(* IEC 61131-3 sources: plc-hackathon-2026/deliver/ME_v3_src (part 2) *)

(* ---- Team_Results.st ---- *)
// Team_Results: YEARLY totals checked by the jury against SimScore.total (tolerance 0.1 %).
// Energies [kWh] and costs [EUR], all LREAL. Updated every simulation step (interval k-1).
VAR_GLOBAL
	E_fne : LREAL;                      // PV production after curtailment
	E_fec : LREAL;                      // fixed consumption
	E_bess_chg : LREAL;                 // battery charge, bus side
	E_bess_dch : LREAL;                 // battery discharge, bus side
	E_ev : LREAL;                       // EV chargers total, bus side
	E_import : LREAL;                   // grid import
	E_export : LREAL;                   // grid export
	E_ev_ch : ARRAY[0..3] OF LREAL;     // per EV charger, bus side
	P_peak : LREAL;                     // [kW] highest monthly peak of the year (info)
	// cost components (spec 4.3)
	C_purchase : LREAL;                 // energy purchase
	C_revenue : LREAL;                  // export revenue (0.9 * price)
	C_grid : LREAL;                     // grid fee
	C_peak : LREAL;                     // peak power cost = sum of 12 monthly values
	C_total : LREAL;                    // purchase - revenue + grid + peak
	// same quantities with the simulator's SimScore.total names
	cost_energy : LREAL;                // purchase - revenue
	cost_grid : LREAL;
	cost_peak : LREAL;
	cost_total : LREAL;
	nLogged : DINT;                     // number of 15-min intervals logged (35040 after the final call)
END_VAR

(* ---- F_AlarmPush.st ---- *)
FUNCTION F_AlarmPush : BOOL
// Push a message into the alarm history (Team_HMI.aAlarmHist, newest at index 0), stamped with simulated time.
VAR_INPUT
	k : DINT;
	sStamp : STRING(20);
	iCode : INT;
	sText : STRING(80);
END_VAR
VAR
	i : INT;
END_VAR
// ---IMPL---
FOR i := 49 TO 1 BY -1 DO
	Team_HMI.aAlarmHist[i] := Team_HMI.aAlarmHist[i - 1];
END_FOR;
Team_HMI.aAlarmHist[0].k := k;
Team_HMI.aAlarmHist[0].sStamp := sStamp;
Team_HMI.aAlarmHist[0].iCode := iCode;
Team_HMI.aAlarmHist[0].sText := sText;
Team_HMI.nAlarms := Team_HMI.nAlarms + 1;
Team_HMI.sLastAlarm := sText;
F_AlarmPush := TRUE;

(* ---- F_BessMaxChg.st ---- *)
FUNCTION F_BessMaxChg : REAL
// Largest bus-side charge power [kW] the simulator accepts at this SoC (same clamp as Sim_Core).
VAR_INPUT
	rSoc : REAL;            // [%] SoC at start of the interval
END_VAR
// ---IMPL---
F_BessMaxChg := LREAL_TO_REAL(MAX(0.0, MIN(REAL_TO_LREAL(SimParam.BESS_MAX_CHG),
	(REAL_TO_LREAL(SimParam.BESS_SOC_MAX) - REAL_TO_LREAL(rSoc)) / 100.0 * REAL_TO_LREAL(SimParam.BESS_CAPACITY)
	/ (REAL_TO_LREAL(SimParam.TS_H) * REAL_TO_LREAL(SimParam.BESS_ETA_CHG)))));

(* ---- F_BessMaxDch.st ---- *)
FUNCTION F_BessMaxDch : REAL
// Largest bus-side discharge power [kW] the simulator accepts at this SoC (same clamp as Sim_Core).
VAR_INPUT
	rSoc : REAL;            // [%] SoC at start of the interval
END_VAR
// ---IMPL---
F_BessMaxDch := LREAL_TO_REAL(MAX(0.0, MIN(REAL_TO_LREAL(SimParam.BESS_MAX_DCH),
	(REAL_TO_LREAL(rSoc) - REAL_TO_LREAL(SimParam.BESS_SOC_MIN)) / 100.0 * REAL_TO_LREAL(SimParam.BESS_CAPACITY)
	* REAL_TO_LREAL(SimParam.BESS_ETA_DCH) / REAL_TO_LREAL(SimParam.TS_H))));

(* ---- F_DayType.st ---- *)
FUNCTION F_DayType : INT
// Day type for load forecasting: 0 = Monday..Friday, 1 = Saturday, 2 = Sunday.
VAR_INPUT
	iWeekday : INT;                     // 1 = Monday .. 7 = Sunday
END_VAR
// ---IMPL---
IF iWeekday = 6 THEN
	F_DayType := 1;
ELSIF iWeekday = 7 THEN
	F_DayType := 2;
ELSE
	F_DayType := 0;
END_IF;

(* ---- F_DtString.st ---- *)
FUNCTION F_DtString : STRING(20)
// DT -> "DD.MM.YYYY HH:MM" (simulated time). Pure calendar arithmetic, no clock access.
VAR_INPUT
	dtIn : DT;
END_VAR
VAR
	udSec : UDINT;
	iDoy : INT;
	iYear : INT;
	iMon : INT;
	iDim : INT;
	xLeap : BOOL;
	uH : USINT;
	uM : USINT;
END_VAR
// ---IMPL---
udSec := DT_TO_UDINT(dtIn);                          // seconds since 1970-01-01
uH := UDINT_TO_USINT((udSec MOD 86400) / 3600);
uM := UDINT_TO_USINT((udSec MOD 3600) / 60);
iDoy := UDINT_TO_INT(udSec / 86400);
iYear := 1970;
xLeap := FALSE;
WHILE iYear < 2200 DO
	xLeap := ((iYear MOD 4) = 0 AND (iYear MOD 100) <> 0) OR ((iYear MOD 400) = 0);
	IF xLeap THEN iDim := 366; ELSE iDim := 365; END_IF;
	IF iDoy < iDim THEN EXIT; END_IF;
	iDoy := iDoy - iDim;
	iYear := iYear + 1;
END_WHILE;
iMon := 1;
WHILE iMon < 12 DO
	CASE iMon OF
		2: IF xLeap THEN iDim := 29; ELSE iDim := 28; END_IF;
		4, 6, 9, 11: iDim := 30;
	ELSE
		iDim := 31;
	END_CASE;
	IF iDoy < iDim THEN EXIT; END_IF;
	iDoy := iDoy - iDim;
	iMon := iMon + 1;
END_WHILE;
F_DtString := CONCAT(CONCAT(CONCAT(F_Pad2(INT_TO_USINT(iDoy + 1)), '.'), CONCAT(F_Pad2(INT_TO_USINT(iMon)), '.')),
	CONCAT(CONCAT(INT_TO_STRING(iYear), ' '), CONCAT(CONCAT(F_Pad2(uH), ':'), F_Pad2(uM))));

(* ---- F_EnergyPrice.st ---- *)
FUNCTION F_EnergyPrice : REAL
// Energy price [EUR/kWh] of interval k for the selected price model (same series the simulator uses).
//   iMode 0 = two-tariff Elektra (per calendar quarter, VT/NT), 1 = day-ahead (Team_Prices.aDA)
VAR_INPUT
	k : DINT;               // interval 0..35039
	iMonth : INT;           // 1..12 of interval k
	xHigh : BOOL;           // VT of interval k (t_sim.tariff_high)
	iMode : INT;            // SimCtrl.price_mode
END_VAR
VAR
	iQ : INT;
END_VAR
// ---IMPL---
IF iMode = 1 THEN
	F_EnergyPrice := Team_Prices.aDA[LIMIT(0, k, 35039)];
ELSE
	iQ := LIMIT(1, (iMonth - 1) / 3 + 1, 4);
	IF xHigh THEN
		F_EnergyPrice := Team_Prices.TT_VT[iQ];
	ELSE
		F_EnergyPrice := Team_Prices.TT_NT[iQ];
	END_IF;
END_IF;

(* ---- F_Pad2.st ---- *)
FUNCTION F_Pad2 : STRING(2)
// Two-digit zero padded number for date/time strings.
VAR_INPUT
	v : USINT;
END_VAR
// ---IMPL---
IF v < 10 THEN
	F_Pad2 := CONCAT('0', USINT_TO_STRING(v));
ELSE
	F_Pad2 := USINT_TO_STRING(v);
END_IF;

(* ---- F_PeakCap.st ---- *)
FUNCTION F_PeakCap : REAL
// Lowest monthly import cap [kW] the battery can hold over the horizon for the given net-load
// forecast (bisection). The battery covers load above the cap and recharges below it.
// Never below rFloor (the peak already paid this month), never above rLimImp.
VAR_INPUT
	h : INT;                            // horizon length
	rE0 : REAL;                         // usable stored energy now [kWh]
	rFloor : REAL;                      // peak already reached this month [kW]
	rLimImp : REAL;                     // import limit [kW]
END_VAR
VAR_IN_OUT
	aLoad : ARRAY[0..191] OF REAL;      // net-load forecast [kW]
END_VAR
VAR
	n : INT;
	i : INT;
	rMid : REAL;
	rLo : REAL;
	rHi : REAL;
	rE : REAL;
	rG : REAL;
	rNeed : REAL;
	rEuse : REAL;
	xOk : BOOL;
END_VAR
// ---IMPL---
rEuse := (SimParam.BESS_SOC_MAX - SimParam.BESS_SOC_MIN) / 100.0 * SimParam.BESS_CAPACITY;
F_PeakCap := rFloor;
rLo := rFloor;
rHi := rLimImp;
FOR n := 0 TO 12 DO
	IF n = 0 THEN
		rMid := rFloor;
	ELSE
		rMid := 0.5 * (rLo + rHi);
	END_IF;
	xOk := TRUE;
	rE := rE0;
	FOR i := 0 TO h - 1 DO
		rG := aLoad[i];
		IF rG > rMid THEN
			rNeed := rG - rMid;
			rE := rE - rNeed * SimParam.TS_H / SimParam.BESS_ETA_DCH;
			IF rNeed > SimParam.BESS_MAX_DCH OR rE < 0.0 THEN
				xOk := FALSE;
				EXIT;
			END_IF;
		ELSE
			rE := rE + MIN(MIN(rMid - rG, SimParam.BESS_MAX_CHG), (rEuse - rE) / (SimParam.TS_H * SimParam.BESS_ETA_CHG))
				* SimParam.TS_H * SimParam.BESS_ETA_CHG;
		END_IF;
	END_FOR;
	IF n = 0 THEN
		IF xOk THEN
			RETURN;                     // the already-paid peak is enough
		END_IF;
	ELSIF xOk THEN
		rHi := rMid;
	ELSE
		rLo := rMid;
	END_IF;
END_FOR;
F_PeakCap := MAX(rFloor, MIN(rLimImp, rHi * Team_Cfg.PLAN_CAPM));

(* ---- F_StageCost.st ---- *)
FUNCTION F_StageCost : REAL
// Cost [EUR] of one 15-min interval, used by FB_Planner.
//   rG >= 0 (import): rG*TS*(price+fee);  rG < 0 (export): -min(-rG, limit)*TS*0.9*price (value >= 0,
//   at negative prices PV is curtailed instead of exporting)
//   + PLAN_PEN * (rGpen - cap) if the (pessimistic) import rGpen would exceed the monthly cap.
VAR_INPUT
	rG : REAL;                          // expected grid power [kW], + import
	rGpen : REAL;                       // pessimistic grid power for the peak penalty [kW]
	rCi : REAL;                         // import price + grid fee [EUR/kWh]
	rCe : REAL;                         // export value [EUR/kWh] (>= 0)
	rT : REAL;                          // import cap [kW]
	rLimExp : REAL;                     // export limit [kW]
END_VAR
// ---IMPL---
IF rG >= 0.0 THEN
	F_StageCost := rG * SimParam.TS_H * rCi;
ELSE
	F_StageCost := -MIN(-rG, rLimExp) * SimParam.TS_H * rCe;
END_IF;
IF rGpen > rT THEN
	F_StageCost := F_StageCost + Team_Cfg.PLAN_PEN * (rGpen - rT);
END_IF;

(* ---- FB_CostLogger.st ---- *)
FUNCTION_BLOCK FB_CostLogger
// Task 3 (spec 4.3): cost logging [EUR] per day / month / year, from the energy of interval k-1
// and the energy price + grid-fee tariff of that same interval.
//   purchase = E_imp * c_en,  revenue = E_exp * 0.9 * c_en,  grid = E_imp * fee(VT/NT)
//   peak (month) = PEAK_PRICE * monthly import peak, year peak = sum of the 12 months
//   day total = purchase - revenue + grid ; month/year total also + peak
// Must be called AFTER FB_EnergyLogger in the same step (uses Team_Log.aMonth[m].P_peak).
VAR_INPUT
	xReset : BOOL;                      // k = 0 (tables are cleared by FB_EnergyLogger)
	xLog : BOOL;                        // log one interval
	iDay : INT;                         // day_of_year of interval k-1
	iMonth : INT;                       // month of interval k-1
	rImp : REAL;                        // EGC_P_import of interval k-1 [kW]
	rExp : REAL;                        // EGC_P_export of interval k-1 [kW]
	rPrice : REAL;                      // energy price of interval k-1 [EUR/kWh]
	xHigh : BOOL;                       // VT tariff of interval k-1 (grid fee)
END_VAR
VAR
	ts : LREAL;
	d : INT;
	m : INT;
	i : INT;
	cBuy : LREAL;
	cRev : LREAL;
	cGrid : LREAL;
	fee : LREAL;
	cPeakYear : LREAL;
END_VAR
// ---IMPL---
IF xLog THEN
	ts := REAL_TO_LREAL(SimParam.TS_H);
	d := LIMIT(0, iDay, 364);
	m := LIMIT(1, iMonth, 12);
	IF xHigh THEN
		fee := REAL_TO_LREAL(SimParam.GRID_VT);
	ELSE
		fee := REAL_TO_LREAL(SimParam.GRID_NT);
	END_IF;
	cBuy := REAL_TO_LREAL(rImp) * ts * REAL_TO_LREAL(rPrice);
	cRev := REAL_TO_LREAL(rExp) * ts * REAL_TO_LREAL(rPrice) * REAL_TO_LREAL(SimParam.EXPORT_FACTOR);
	cGrid := REAL_TO_LREAL(rImp) * ts * fee;

	// day (no peak component)
	Team_Log.aDay[d].C_purchase := Team_Log.aDay[d].C_purchase + cBuy;
	Team_Log.aDay[d].C_revenue := Team_Log.aDay[d].C_revenue + cRev;
	Team_Log.aDay[d].C_grid := Team_Log.aDay[d].C_grid + cGrid;
	Team_Log.aDay[d].C_total := Team_Log.aDay[d].C_purchase - Team_Log.aDay[d].C_revenue + Team_Log.aDay[d].C_grid;
	// month (peak known so far in this month)
	Team_Log.aMonth[m].C_purchase := Team_Log.aMonth[m].C_purchase + cBuy;
	Team_Log.aMonth[m].C_revenue := Team_Log.aMonth[m].C_revenue + cRev;
	Team_Log.aMonth[m].C_grid := Team_Log.aMonth[m].C_grid + cGrid;
	Team_Log.aMonth[m].C_peak := Team_Log.aMonth[m].P_peak * REAL_TO_LREAL(SimParam.PEAK_PRICE);
	Team_Log.aMonth[m].C_total := Team_Log.aMonth[m].C_purchase - Team_Log.aMonth[m].C_revenue
		+ Team_Log.aMonth[m].C_grid + Team_Log.aMonth[m].C_peak;
	// year
	Team_Log.stYear.C_purchase := Team_Log.stYear.C_purchase + cBuy;
	Team_Log.stYear.C_revenue := Team_Log.stYear.C_revenue + cRev;
	Team_Log.stYear.C_grid := Team_Log.stYear.C_grid + cGrid;
	cPeakYear := 0.0;
	FOR i := 1 TO 12 DO
		cPeakYear := cPeakYear + Team_Log.aMonth[i].C_peak;
	END_FOR;
	Team_Log.stYear.C_peak := cPeakYear;
	Team_Log.stYear.C_total := Team_Log.stYear.C_purchase - Team_Log.stYear.C_revenue
		+ Team_Log.stYear.C_grid + Team_Log.stYear.C_peak;
END_IF;

IF xReset OR xLog THEN
	Team_Results.C_purchase := Team_Log.stYear.C_purchase;
	Team_Results.C_revenue := Team_Log.stYear.C_revenue;
	Team_Results.C_grid := Team_Log.stYear.C_grid;
	Team_Results.C_peak := Team_Log.stYear.C_peak;
	Team_Results.C_total := Team_Log.stYear.C_total;
	// simulator (SimScore.total) naming
	Team_Results.cost_energy := Team_Log.stYear.C_purchase - Team_Log.stYear.C_revenue;
	Team_Results.cost_grid := Team_Log.stYear.C_grid;
	Team_Results.cost_peak := Team_Log.stYear.C_peak;
	Team_Results.cost_total := Team_Log.stYear.C_total;
END_IF;

(* ---- FB_EnergyLogger.st ---- *)
FUNCTION_BLOCK FB_EnergyLogger
// Task 2 (spec 4.2): energy logging [kWh] per day / month / year + monthly import peak [kW].
// Called once per NEW simulation step k with the ACTUAL powers of interval k-1 (*_act, EGC_*),
// the fixed consumption remembered from the previous call and the day/month of interval k-1.
// E = P * TS_H, accumulated in LREAL into Team_Log (aDay, aMonth, stYear) and Team_Results.
VAR_INPUT
	xReset : BOOL;                      // k = 0: clear all tables
	xLog : BOOL;                        // log one interval
	iDay : INT;                         // day_of_year of interval k-1 (0..364)
	iMonth : INT;                       // month of interval k-1 (1..12)
	rFne : REAL;                        // FNE_P_act
	rFec : REAL;                        // FEC_P_fix of interval k-1 (remembered)
	rChg : REAL;                        // BESS_P_charge_act
	rDch : REAL;                        // BESS_P_discharge_act
	aEv : ARRAY[0..3] OF REAL;          // EV[j].P_charge_act
	rImp : REAL;                        // EGC_P_import
	rExp : REAL;                        // EGC_P_export
END_VAR
VAR
	stZero : typeTeamAgg;               // never written -> all zero
	ts : LREAL;
	d : INT;
	m : INT;
	j : INT;
	i : INT;
	eEv : LREAL;
END_VAR
// ---IMPL---
IF xReset THEN
	FOR i := 0 TO 364 DO
		Team_Log.aDay[i] := stZero;
	END_FOR;
	FOR i := 1 TO 12 DO
		Team_Log.aMonth[i] := stZero;
	END_FOR;
	Team_Log.stYear := stZero;
END_IF;

IF xLog THEN
	ts := REAL_TO_LREAL(SimParam.TS_H);
	d := LIMIT(0, iDay, 364);
	m := LIMIT(1, iMonth, 12);
	// day
	Team_Log.aDay[d].E_fne := Team_Log.aDay[d].E_fne + REAL_TO_LREAL(rFne) * ts;
	Team_Log.aDay[d].E_fec := Team_Log.aDay[d].E_fec + REAL_TO_LREAL(rFec) * ts;
	Team_Log.aDay[d].E_bess_chg := Team_Log.aDay[d].E_bess_chg + REAL_TO_LREAL(rChg) * ts;
	Team_Log.aDay[d].E_bess_dch := Team_Log.aDay[d].E_bess_dch + REAL_TO_LREAL(rDch) * ts;
	Team_Log.aDay[d].E_import := Team_Log.aDay[d].E_import + REAL_TO_LREAL(rImp) * ts;
	Team_Log.aDay[d].E_export := Team_Log.aDay[d].E_export + REAL_TO_LREAL(rExp) * ts;
	Team_Log.aDay[d].P_peak := MAX(Team_Log.aDay[d].P_peak, REAL_TO_LREAL(rImp));
	// month
	Team_Log.aMonth[m].E_fne := Team_Log.aMonth[m].E_fne + REAL_TO_LREAL(rFne) * ts;
	Team_Log.aMonth[m].E_fec := Team_Log.aMonth[m].E_fec + REAL_TO_LREAL(rFec) * ts;
	Team_Log.aMonth[m].E_bess_chg := Team_Log.aMonth[m].E_bess_chg + REAL_TO_LREAL(rChg) * ts;
	Team_Log.aMonth[m].E_bess_dch := Team_Log.aMonth[m].E_bess_dch + REAL_TO_LREAL(rDch) * ts;
	Team_Log.aMonth[m].E_import := Team_Log.aMonth[m].E_import + REAL_TO_LREAL(rImp) * ts;
	Team_Log.aMonth[m].E_export := Team_Log.aMonth[m].E_export + REAL_TO_LREAL(rExp) * ts;
	Team_Log.aMonth[m].P_peak := MAX(Team_Log.aMonth[m].P_peak, REAL_TO_LREAL(rImp));
	// year
	Team_Log.stYear.E_fne := Team_Log.stYear.E_fne + REAL_TO_LREAL(rFne) * ts;
	Team_Log.stYear.E_fec := Team_Log.stYear.E_fec + REAL_TO_LREAL(rFec) * ts;
	Team_Log.stYear.E_bess_chg := Team_Log.stYear.E_bess_chg + REAL_TO_LREAL(rChg) * ts;
	Team_Log.stYear.E_bess_dch := Team_Log.stYear.E_bess_dch + REAL_TO_LREAL(rDch) * ts;
	Team_Log.stYear.E_import := Team_Log.stYear.E_import + REAL_TO_LREAL(rImp) * ts;
	Team_Log.stYear.E_export := Team_Log.stYear.E_export + REAL_TO_LREAL(rExp) * ts;
	Team_Log.stYear.P_peak := MAX(Team_Log.stYear.P_peak, REAL_TO_LREAL(rImp));
	// EV per charger and total
	FOR j := 0 TO 3 DO
		eEv := REAL_TO_LREAL(aEv[j]) * ts;
		Team_Log.aDay[d].E_ev_ch[j] := Team_Log.aDay[d].E_ev_ch[j] + eEv;
		Team_Log.aDay[d].E_ev := Team_Log.aDay[d].E_ev + eEv;
		Team_Log.aMonth[m].E_ev_ch[j] := Team_Log.aMonth[m].E_ev_ch[j] + eEv;
		Team_Log.aMonth[m].E_ev := Team_Log.aMonth[m].E_ev + eEv;
		Team_Log.stYear.E_ev_ch[j] := Team_Log.stYear.E_ev_ch[j] + eEv;
		Team_Log.stYear.E_ev := Team_Log.stYear.E_ev + eEv;
	END_FOR;
END_IF;

IF xReset OR xLog THEN
	// publish yearly energies (names required by spec 4.2)
	Team_Results.E_fne := Team_Log.stYear.E_fne;
	Team_Results.E_fec := Team_Log.stYear.E_fec;
	Team_Results.E_bess_chg := Team_Log.stYear.E_bess_chg;
	Team_Results.E_bess_dch := Team_Log.stYear.E_bess_dch;
	Team_Results.E_ev := Team_Log.stYear.E_ev;
	Team_Results.E_import := Team_Log.stYear.E_import;
	Team_Results.E_export := Team_Log.stYear.E_export;
	Team_Results.E_ev_ch := Team_Log.stYear.E_ev_ch;
	Team_Results.P_peak := Team_Log.stYear.P_peak;
	IF xReset THEN
		Team_Results.nLogged := 0;
	END_IF;
	IF xLog THEN
		Team_Results.nLogged := Team_Results.nLogged + 1;
	END_IF;
END_IF;

(* ---- FB_Forecast.st ---- *)
FUNCTION_BLOCK FB_Forecast
// Forecast of the next h intervals (allowed by spec 4.1: estimates from PAST data only).
//   FEC: exponential moving average per day type (Mon-Fri / Sat / Sun) and quarter-hour,
//        plus the mean absolute deviation (sigma) per day type and quarter-hour.
//   PV : exponential moving average per quarter-hour (all days).
//   Intraday correction: ratio actual / profile over the last FC_CORR_W intervals scales the
//        profile forecast, fading out with time constant FC_CORR_TAU (cloudy day, busy day ...).
//   VT : tariff window learned from the last observed day.
//   EV : connected vehicles charged as soon as possible with their remaining energy.
// Interval i = 0 is the current interval k and uses the ACTUAL simOut values.
// Outputs: aNet = expected net load, aNetHi = pessimistic net load (for the peak cap):
//          + rKsig * sigma(FEC) + (1 - PLAN_PVF) * PV forecast.
// Learned profiles live in this FB only (built online from simOut, nothing is embedded).
VAR_INPUT
	xReset : BOOL;                      // k = 0: forget all learned profiles
	xUpdate : BOOL;                     // new step: learn from the current interval
	k : DINT;                           // current step
	iQh : INT;                          // qh_of_day of k
	iWeekday : INT;                     // 1 = Mon .. 7 = Sun of k
	rFec : REAL;                        // FEC_P_fix of k
	rPv : REAL;                         // FNE_output_power of k
	xVt : BOOL;                         // tariff_high of k
	aEvRem : ARRAY[0..3] OF REAL;       // EV remaining energy [kWh] (0 if not connected)
	aEvSteps : ARRAY[0..3] OF DINT;     // EV steps to departure
	iH : INT;                           // horizon length (1..192)
	rKsig : REAL;                       // pessimistic load = expected + rKsig * sigma
END_VAR
VAR_IN_OUT
	aNet : ARRAY[0..191] OF REAL;       // expected net load fec + ev - pv [kW]
	aNetHi : ARRAY[0..191] OF REAL;     // pessimistic net load [kW]
	aVtF : ARRAY[0..191] OF BOOL;       // forecast VT
END_VAR
VAR
	aFec : ARRAY[0..2, 0..95] OF REAL;  // learned FEC profile per day type
	aSig : ARRAY[0..2, 0..95] OF REAL;  // learned mean abs deviation of FEC
	aFecOk : ARRAY[0..2, 0..95] OF BOOL;
	aPv : ARRAY[0..95] OF REAL;         // learned PV profile
	aPvOk : ARRAY[0..95] OF BOOL;
	aVt : ARRAY[0..95] OF BOOL;         // last observed VT window
	aHf : ARRAY[0..15] OF REAL;         // recent actual FEC
	aHfP : ARRAY[0..15] OF REAL;        // profile value for it (before update)
	aHp : ARRAY[0..15] OF REAL;         // recent actual PV
	aHpP : ARRAY[0..15] OF REAL;        // profile value for it
	nHist : INT;                        // valid entries in the ring
	iHead : INT;                        // next write index
	rCorrF : REAL := 1.0;               // FEC intraday ratio
	rCorrP : REAL := 1.0;               // PV intraday ratio
	rFecMax : REAL;                     // highest FEC seen since reset (cold-start fallback)
	aEvR : ARRAY[0..3] OF REAL;
	i : INT;
	j : INT;
	q : INT;
	dtp : INT;
	wd : INT;
	kk : DINT;
	rF : REAL;
	rP : REAL;
	rS : REAL;
	rEv : REAL;
	pe : REAL;
	rA : REAL;
	rB : REAL;
	rA2 : REAL;
	rB2 : REAL;
	rDecay : REAL;
	rPrevF : REAL;
	rPrevP : REAL;
END_VAR
// ---IMPL---
IF xReset THEN
	FOR q := 0 TO 95 DO
		FOR dtp := 0 TO 2 DO
			aFec[dtp, q] := 0.0;
			aSig[dtp, q] := 0.0;
			aFecOk[dtp, q] := FALSE;
		END_FOR;
		aPv[q] := 0.0;
		aPvOk[q] := FALSE;
		aVt[q] := FALSE;
	END_FOR;
	nHist := 0;
	iHead := 0;
	rFecMax := 0.0;
	rCorrF := 1.0;
	rCorrP := 1.0;
END_IF;

// ---- learn from the current interval ----
IF xUpdate THEN
	q := LIMIT(0, iQh, 95);
	dtp := F_DayType(iWeekday);
	rFecMax := MAX(rFecMax, rFec);
	// profile values before the update (for the intraday ratio)
	IF aFecOk[dtp, q] THEN rPrevF := aFec[dtp, q]; ELSE rPrevF := rFec; END_IF;
	IF aPvOk[q] THEN rPrevP := aPv[q]; ELSE rPrevP := rPv; END_IF;
	IF aFecOk[dtp, q] THEN
		aSig[dtp, q] := aSig[dtp, q] + Team_Cfg.FC_ALPHA_SIG * (ABS(rFec - aFec[dtp, q]) - aSig[dtp, q]);
		aFec[dtp, q] := aFec[dtp, q] + Team_Cfg.FC_ALPHA_FEC * (rFec - aFec[dtp, q]);
	ELSE
		aFec[dtp, q] := rFec;
		aFecOk[dtp, q] := TRUE;
	END_IF;
	IF aPvOk[q] THEN
		aPv[q] := aPv[q] + Team_Cfg.FC_ALPHA_PV * (rPv - aPv[q]);
	ELSE
		aPv[q] := rPv;
		aPvOk[q] := TRUE;
	END_IF;
	aVt[q] := xVt;
	// intraday correction ratios over the last FC_CORR_W intervals
	IF Team_Cfg.FC_CORR_W > 0 THEN
		aHf[iHead] := rFec;
		aHfP[iHead] := rPrevF;
		aHp[iHead] := rPv;
		aHpP[iHead] := rPrevP;
		iHead := (iHead + 1) MOD 16;
		nHist := MIN(nHist + 1, LIMIT(1, Team_Cfg.FC_CORR_W, 16));
		rA := 0.0; rB := 0.0; rA2 := 0.0; rB2 := 0.0;
		FOR j := 1 TO nHist DO
			i := (iHead - j + 16) MOD 16;
			rA := rA + aHf[i];
			rB := rB + aHfP[i];
			rA2 := rA2 + aHp[i];
			rB2 := rB2 + aHpP[i];
		END_FOR;
		IF Team_Cfg.FC_CORR_FEC AND rB > 10.0 THEN
			rCorrF := LIMIT(0.5, rA / rB, 1.5);
		ELSE
			rCorrF := 1.0;
		END_IF;
		IF Team_Cfg.FC_CORR_PV AND rB2 > 20.0 THEN
			rCorrP := LIMIT(0.2, rA2 / rB2, 1.5);
		ELSE
			rCorrP := 1.0;
		END_IF;
	END_IF;
END_IF;

// ---- horizon ----
FOR j := 0 TO 3 DO
	aEvR[j] := aEvRem[j];
END_FOR;
FOR i := 0 TO LIMIT(1, iH, 192) - 1 DO
	kk := k + i;
	q := DINT_TO_INT(kk MOD 96);
	rS := 0.0;
	IF i = 0 THEN
		rF := rFec;
		rP := rPv;
		aVtF[i] := xVt;
	ELSE
		wd := DINT_TO_INT((INT_TO_DINT(iWeekday) - 1 + (kk / 96) - (k / 96)) MOD 7) + 1;
		dtp := F_DayType(wd);
		IF aFecOk[dtp, q] THEN
			rF := aFec[dtp, q];
			rS := aSig[dtp, q];
		ELSIF aFecOk[0, q] THEN
			rF := aFec[0, q];
		ELSE
			rF := rFecMax;              // nothing learned yet (first day): assume the highest load seen so far
		END_IF;
		rP := aPv[q];
		IF Team_Cfg.FC_CORR_W > 0 THEN
			rDecay := EXP(-INT_TO_REAL(i) / Team_Cfg.FC_CORR_TAU);
			rF := rF * (1.0 + (rCorrF - 1.0) * rDecay);
			rP := rP * (1.0 + (rCorrP - 1.0) * rDecay);
		END_IF;
		aVtF[i] := aVt[q];
	END_IF;
	rEv := 0.0;
	FOR j := 0 TO 3 DO
		IF aEvR[j] > 0.000001 AND i < aEvSteps[j] THEN
			pe := MIN(SimParam.EV_MAX_CHARGE, aEvR[j] / (SimParam.TS_H * SimParam.EV_ETA));
			aEvR[j] := aEvR[j] - pe * SimParam.TS_H * SimParam.EV_ETA;
			rEv := rEv + pe;
		END_IF;
	END_FOR;
	aNet[i] := rF + rEv - rP;
	IF i = 0 THEN
		aNetHi[i] := aNet[i];
	ELSE
		aNetHi[i] := aNet[i] + rKsig * rS + (1.0 - Team_Cfg.PLAN_PVF) * rP;
	END_IF;
END_FOR;

(* ---- FB_GridGuard.st ---- *)
FUNCTION_BLOCK FB_GridGuard
// Grid-connection protection (spec 2.5 / 4.1, mandatory). Always the LAST stage before simCmd.
// Predicts the grid power of the CURRENT interval from the bus balance
//     P_grid = P_fec - P_fne + sum(P_ev) - P_bess      (P_bess: + discharge, - charge)
// using the values the simulator will actually realise (same clamps as Sim_Core: SoC limits,
// EV remaining energy, PV availability), and corrects the requested setpoints so that
//     P_grid <= EGC_MAX_IMPORT - margin   and   -P_grid <= EGC_MAX_EXPORT - margin.
// Import side: 1) drop voluntary curtailment, 2) more BESS discharge, 3) shed EV power (most slack first).
// Export side: 1) less discharge / more BESS charge, 2) curtail PV (safer than relying on the battery).
VAR_INPUT
	rFec : REAL;                        // fixed consumption of interval k [kW]
	rFneAvail : REAL;                   // available PV of interval k [kW]
	rBcMax : REAL;                      // feasible BESS charge [kW] (F_BessMaxChg)
	rBdMax : REAL;                      // feasible BESS discharge [kW] (F_BessMaxDch)
	aEvMax : ARRAY[0..3] OF REAL;       // feasible EV power per charger [kW] (0 if not connected)
	aEvSlack : ARRAY[0..3] OF REAL;     // EV scheduling slack [steps], bigger = shed first
	rPbReq : REAL;                      // requested BESS power, + discharge / - charge
	aEvReq : ARRAY[0..3] OF REAL;       // requested EV powers
	xCurtReq : BOOL;                    // strategy wants curtailment (e.g. negative price)
	rCurtReq : REAL;                    // requested PV limit [kW]
END_VAR
VAR_OUTPUT
	rPb : REAL;                         // final BESS power, + discharge / - charge
	aEv : ARRAY[0..3] OF REAL;          // final EV powers
	xCurt : BOOL;                       // final curtailment enable
	rCurt : REAL;                       // final PV limit [kW]
	rFne : REAL;                        // expected PV after curtailment
	rGridPred : REAL;                   // predicted grid power, + import / - export
	xEvShed : BOOL;                     // EV power reduced by the guard
	xExpCurt : BOOL;                    // PV curtailed by the guard for export protection
	xImpFail : BOOL;                    // import limit cannot be held (should never happen)
END_VAR
VAR
	limImp : REAL;
	limExp : REAL;
	sumEv : REAL;
	pg : REAL;
	d : REAL;
	j : INT;
	jSel : INT;
	n : INT;
	rBest : REAL;
END_VAR
// ---IMPL---
limImp := SimParam.EGC_MAX_IMPORT - Team_Cfg.GRID_MARGIN_IMP;
limExp := SimParam.EGC_MAX_EXPORT - Team_Cfg.GRID_MARGIN_EXP;
xEvShed := FALSE;
xExpCurt := FALSE;
xImpFail := FALSE;

// 1. clamp requests to what the simulator will realise
rPb := LIMIT(-rBcMax, rPbReq, rBdMax);
sumEv := 0.0;
FOR j := 0 TO 3 DO
	aEv[j] := LIMIT(0.0, aEvReq[j], aEvMax[j]);
	sumEv := sumEv + aEv[j];
END_FOR;
IF xCurtReq THEN
	rFne := MIN(rFneAvail, MAX(0.0, rCurtReq));
ELSE
	rFne := rFneAvail;
END_IF;
pg := rFec - rFne + sumEv - rPb;

// 2. import protection
IF pg > limImp THEN
	// 2a. give back voluntarily curtailed PV
	d := MIN(pg - limImp, rFneAvail - rFne);
	IF d > 0.0 THEN
		rFne := rFne + d;
		pg := pg - d;
	END_IF;
	// 2b. more discharge
	d := MIN(pg - limImp, rBdMax - rPb);
	IF d > 0.0 THEN
		rPb := rPb + d;
		pg := pg - d;
	END_IF;
	// 2c. shed EV power, charger with the largest slack first
	n := 0;
	WHILE pg > limImp AND n < 4 DO
		jSel := -1;
		rBest := -1.0E30;
		FOR j := 0 TO 3 DO
			IF aEv[j] > 0.0 AND aEvSlack[j] > rBest THEN
				rBest := aEvSlack[j];
				jSel := j;
			END_IF;
		END_FOR;
		IF jSel < 0 THEN
			EXIT;
		END_IF;
		d := MIN(pg - limImp, aEv[jSel]);
		aEv[jSel] := aEv[jSel] - d;
		sumEv := sumEv - d;
		pg := pg - d;
		xEvShed := TRUE;
		n := n + 1;
	END_WHILE;
	xImpFail := pg > limImp;
END_IF;

// 3. export protection
IF pg < -limExp THEN
	// 3a. less discharge / more charge
	d := MIN(-limExp - pg, rPb + rBcMax);
	IF d > 0.0 THEN
		rPb := rPb - d;
		pg := pg + d;
	END_IF;
	// 3b. curtail PV
	IF pg < -limExp THEN
		rFne := MAX(0.0, rFne - (-limExp - pg));
		xExpCurt := TRUE;
	END_IF;
END_IF;

// 4. outputs
xCurt := rFne < rFneAvail - 0.0001;
IF xCurt THEN
	rCurt := rFne;
ELSE
	rCurt := 0.0;
	rFne := rFneAvail;
END_IF;
sumEv := 0.0;
FOR j := 0 TO 3 DO
	sumEv := sumEv + aEv[j];
END_FOR;
rGridPred := rFec - rFne + sumEv - rPb;

(* ---- FB_HmiUpdate.st ---- *)
FUNCTION_BLOCK FB_HmiUpdate
// Fills Team_HMI for the HMI: simulated date/time, progress, requested vs actual flows, SoC, EVs,
// table selections, 24 h trends (96 samples, simulated time) and the alarm/message history.
// Trends and alarms advance only on a NEW simulation step -> independent of the PLC cycle time.
VAR_INPUT
	xNewStep : BOOL;                    // first call of a new step k
	xReset : BOOL;                      // k = 0 after reset
	stOut : typeSimOut;                 // simulator outputs (copy of simOut)
	stCmd : typeSimCmd;                 // commands issued for interval k
	rPbCmd : REAL;                      // final BESS setpoint, + discharge / - charge
	rFneExp : REAL;                     // expected PV after curtailment
	rGridPred : REAL;                   // predicted grid power interval k
	rFecPrev : REAL;                    // fixed consumption interval k-1
	rPrice : REAL;                      // energy price interval k
	rPricePrev : REAL;                  // energy price interval k-1
	aEvSteps : ARRAY[0..3] OF DINT;     // steps to departure
	aEvLast : ARRAY[0..3] OF REAL;      // actual EV power of interval k-1 (corrected for departures)
	rPeakMonth : REAL;                  // running monthly import peak
	rPeakTarget : REAL;                 // controller import cap
	xEvShed : BOOL;                     // guard flags of this step
	xExpCurt : BOOL;
	xImpFail : BOOL;
END_VAR
VAR
	i : INT;
	j : INT;
	iSel : INT;
	iFirst : INT;
	rGridPredLast : REAL;               // prediction made for the previous interval
	xHavePred : BOOL;
	aPrevConn : ARRAY[0..3] OF BOOL;
	aPrevRemain : ARRAY[0..3] OF REAL;
	aPrevDepK : ARRAY[0..3] OF DINT;
	xPrevImpOv : BOOL;
	xPrevExpOv : BOOL;
	xPrevTrip : BOOL;
	xPrevFin : BOOL;
	xPrevShed : BOOL;
	xPrevCurt : BOOL;
	xPrevFail : BOOL;
	rUnmet : REAL;
	aDim : ARRAY[1..12] OF INT := [31, 28, 31, 30, 31, 30, 31, 31, 30, 31, 30, 31];
	stZero : typeTeamAgg;
	kNow : DINT;
END_VAR
// ---IMPL---
kNow := stOut.t_sim.k;
Team_HMI.nCalls := Team_HMI.nCalls + 1;

// ---------------- reset (k = 0) ----------------
IF xReset THEN
	FOR i := 0 TO 95 DO
		Team_HMI.aTrFne[i] := 0.0;
		Team_HMI.aTrFec[i] := 0.0;
		Team_HMI.aTrGrid[i] := 0.0;
		Team_HMI.aTrBess[i] := 0.0;
		Team_HMI.aTrEv[i] := 0.0;
		Team_HMI.aTrSoc[i] := 0.0;
		Team_HMI.aTrPrice[i] := 0.0;
	END_FOR;
	FOR i := 0 TO 49 DO
		Team_HMI.aAlarmHist[i].k := 0;
		Team_HMI.aAlarmHist[i].sStamp := '';
		Team_HMI.aAlarmHist[i].iCode := 0;
		Team_HMI.aAlarmHist[i].sText := '';
	END_FOR;
	Team_HMI.nAlarms := 0;
	Team_HMI.sLastAlarm := '';
	Team_HMI.nSteps := 0;
	Team_HMI.nGuardEv := 0;
	Team_HMI.nGuardCurt := 0;
	Team_HMI.nGuardFail := 0;
	Team_HMI.nBothEnables := 0;
	Team_HMI.rEvUnmetSum := 0.0;
	Team_HMI.rGridPredErr := 0.0;
	Team_HMI.rGridPredErrMax := 0.0;
	Team_HMI.xAlmEvUnmet := FALSE;
	xHavePred := FALSE;
	xPrevImpOv := FALSE;
	xPrevExpOv := FALSE;
	xPrevTrip := FALSE;
	xPrevFin := FALSE;
	xPrevShed := FALSE;
	xPrevCurt := FALSE;
	xPrevFail := FALSE;
	FOR j := 0 TO 3 DO
		aPrevConn[j] := FALSE;
	END_FOR;
END_IF;

// ---------------- status / header (every call) ----------------
Team_HMI.sDateTime := F_DtString(stOut.t_sim.stamp);
Team_HMI.k := kNow;
Team_HMI.rProgressPct := DINT_TO_REAL(kNow) * 100.0 / DINT_TO_REAL(Team_Cfg.N_STEPS);
Team_HMI.xTariffHigh := stOut.t_sim.tariff_high;
IF stOut.t_sim.tariff_high THEN
	Team_HMI.sTariff := 'VT';
	Team_HMI.rGridFee := SimParam.GRID_VT;
ELSE
	Team_HMI.sTariff := 'NT';
	Team_HMI.rGridFee := SimParam.GRID_NT;
END_IF;
IF SimCtrl.price_mode = 1 THEN
	Team_HMI.sPriceMode := 'Dan-unaprijed';
ELSE
	Team_HMI.sPriceMode := 'Dvotarifni (HEP)';
END_IF;
Team_HMI.rPrice := rPrice;

// requested (interval k)
Team_HMI.rFneAvail := stOut.FNE_output_power;
Team_HMI.rFneExpected := rFneExp;
Team_HMI.xCurtActive := stCmd.FNE_enable_curtail;
Team_HMI.rCurtValue := stCmd.FNE_curtail_value;
Team_HMI.rFec := stOut.FEC_P_fix;
Team_HMI.rFecPrev := rFecPrev;
Team_HMI.rBessReq := rPbCmd;
Team_HMI.rBessChgReq := SEL(stCmd.BESS_enable_charge, 0.0, stCmd.BESS_P_charge);
Team_HMI.rBessDchReq := SEL(stCmd.BESS_enable_discharge, 0.0, stCmd.BESS_P_discharge);
Team_HMI.rGridPred := rGridPred;
Team_HMI.rEvReqSum := 0.0;
Team_HMI.rEvActSum := 0.0;
FOR j := 0 TO 3 DO
	Team_HMI.aEvReq[j] := stCmd.EV[j].P_charge;
	Team_HMI.aEvAct[j] := aEvLast[j];
	Team_HMI.rEvReqSum := Team_HMI.rEvReqSum + stCmd.EV[j].P_charge;
	Team_HMI.rEvActSum := Team_HMI.rEvActSum + aEvLast[j];
	Team_HMI.aEvConnected[j] := stOut.EV[j].connected;
	IF stOut.EV[j].connected THEN
		Team_HMI.aEvDeparture[j] := F_DtString(stOut.EV[j].planned_departure);
	ELSE
		Team_HMI.aEvDeparture[j] := '';
	END_IF;
	Team_HMI.aEvRemaining[j] := stOut.EV[j].energy_required;
	Team_HMI.aEvDelivered[j] := stOut.EV[j].energy_delivered;
	Team_HMI.aEvStepsLeft[j] := aEvSteps[j];
END_FOR;
// actual (interval k-1)
Team_HMI.rFneAct := stOut.FNE_P_act;
Team_HMI.rBessChgAct := stOut.BESS_P_charge_act;
Team_HMI.rBessDchAct := stOut.BESS_P_discharge_act;
Team_HMI.rBessAct := stOut.BESS_P_discharge_act - stOut.BESS_P_charge_act;
Team_HMI.rImportAct := stOut.EGC_P_import;
Team_HMI.rExportAct := stOut.EGC_P_export;
// battery
Team_HMI.rSoc := stOut.BESS_SoC;
Team_HMI.rSocMin := SimParam.BESS_SOC_MIN;
Team_HMI.rSocMax := SimParam.BESS_SOC_MAX;
IF rPbCmd > Team_Cfg.P_EPS THEN
	Team_HMI.sBessDir := 'PRAZNJENJE';
ELSIF rPbCmd < -Team_Cfg.P_EPS THEN
	Team_HMI.sBessDir := 'PUNJENJE';
ELSE
	Team_HMI.sBessDir := 'MIROVANJE';
END_IF;
Team_HMI.rPeakMonth := rPeakMonth;
Team_HMI.rPeakTarget := rPeakTarget;
IF stCmd.BESS_enable_charge AND stCmd.BESS_enable_discharge THEN
	Team_HMI.nBothEnables := Team_HMI.nBothEnables + 1;
END_IF;

// ---------------- table selection (HMI writes iSelDay / iSelMonth) ----------------
iSel := LIMIT(0, Team_HMI.iSelDay, 364);
Team_HMI.stSelDay := Team_Log.aDay[iSel];
iSel := LIMIT(1, Team_HMI.iSelMonth, 12);
Team_HMI.stSelMonth := Team_Log.aMonth[iSel];
Team_HMI.iSelMonthDays := aDim[iSel];
iFirst := 0;
FOR i := 1 TO iSel - 1 DO
	iFirst := iFirst + aDim[i];
END_FOR;
FOR i := 1 TO 31 DO
	IF i <= aDim[iSel] THEN
		Team_HMI.aSelMonthDays[i] := Team_Log.aDay[iFirst + i - 1];
	ELSE
		Team_HMI.aSelMonthDays[i] := stZero;
	END_IF;
END_FOR;

// ---------------- once per new step: trends, prediction check, alarms ----------------
IF xNewStep THEN
	Team_HMI.nSteps := Team_HMI.nSteps + 1;
	IF kNow > 0 THEN
		// trends: shift left, newest (interval k-1) at index 95
		FOR i := 0 TO 94 DO
			Team_HMI.aTrFne[i] := Team_HMI.aTrFne[i + 1];
			Team_HMI.aTrFec[i] := Team_HMI.aTrFec[i + 1];
			Team_HMI.aTrGrid[i] := Team_HMI.aTrGrid[i + 1];
			Team_HMI.aTrBess[i] := Team_HMI.aTrBess[i + 1];
			Team_HMI.aTrEv[i] := Team_HMI.aTrEv[i + 1];
			Team_HMI.aTrSoc[i] := Team_HMI.aTrSoc[i + 1];
			Team_HMI.aTrPrice[i] := Team_HMI.aTrPrice[i + 1];
		END_FOR;
		Team_HMI.aTrFne[95] := stOut.FNE_P_act;
		Team_HMI.aTrFec[95] := rFecPrev;
		Team_HMI.aTrGrid[95] := stOut.EGC_P_import - stOut.EGC_P_export;
		Team_HMI.aTrBess[95] := stOut.BESS_P_discharge_act - stOut.BESS_P_charge_act;
		Team_HMI.aTrEv[95] := Team_HMI.rEvActSum;
		Team_HMI.aTrSoc[95] := stOut.BESS_SoC;
		Team_HMI.aTrPrice[95] := rPricePrev;
		// grid prediction quality (prediction for k-1 vs measurement of k-1)
		IF xHavePred THEN
			Team_HMI.rGridPredErr := ABS(rGridPredLast - (stOut.EGC_P_import - stOut.EGC_P_export));
			Team_HMI.rGridPredErrMax := MAX(Team_HMI.rGridPredErrMax, Team_HMI.rGridPredErr);
		END_IF;
		// EV departures with undelivered energy
		FOR j := 0 TO 3 DO
			IF aPrevConn[j] AND kNow >= aPrevDepK[j] THEN
				rUnmet := aPrevRemain[j] - aEvLast[j] * SimParam.TS_H * SimParam.EV_ETA;
				IF rUnmet > 0.01 THEN
					Team_HMI.xAlmEvUnmet := TRUE;
					Team_HMI.rEvUnmetSum := Team_HMI.rEvUnmetSum + rUnmet;
					F_AlarmPush(k := kNow, sStamp := Team_HMI.sDateTime, iCode := 5,
						sText := CONCAT(CONCAT('EV punjac ', INT_TO_STRING(j + 1)),
							CONCAT(': vozilo otislo, nepredano kWh = ', REAL_TO_STRING(rUnmet))));
				END_IF;
			END_IF;
		END_FOR;
	END_IF;
	// overload flags of the previous interval (also show as active alarms)
	Team_HMI.xAlmImport := stOut.EGC_overload_import;
	Team_HMI.xAlmExport := stOut.EGC_overload_export;
	IF stOut.EGC_overload_import AND NOT xPrevImpOv THEN
		F_AlarmPush(k := kNow, sStamp := Team_HMI.sDateTime, iCode := 1, sText := 'Prekoracenje uvoza iz mreze (EGC overload import)');
	END_IF;
	IF stOut.EGC_overload_export AND NOT xPrevExpOv THEN
		F_AlarmPush(k := kNow, sStamp := Team_HMI.sDateTime, iCode := 2, sText := 'Prekoracenje izvoza u mrezu (EGC overload export)');
	END_IF;
	xPrevImpOv := stOut.EGC_overload_import;
	xPrevExpOv := stOut.EGC_overload_export;
	// guard interventions (rising edge -> message)
	Team_HMI.xAlmGuardEv := xEvShed;
	Team_HMI.xAlmGuardCurt := xExpCurt;
	Team_HMI.xAlmGuardFail := xImpFail;
	IF xEvShed THEN Team_HMI.nGuardEv := Team_HMI.nGuardEv + 1; END_IF;
	IF xExpCurt THEN Team_HMI.nGuardCurt := Team_HMI.nGuardCurt + 1; END_IF;
	IF xImpFail THEN Team_HMI.nGuardFail := Team_HMI.nGuardFail + 1; END_IF;
	IF xEvShed AND NOT xPrevShed THEN
		F_AlarmPush(k := kNow, sStamp := Team_HMI.sDateTime, iCode := 6, sText := 'Zastita prikljucka: smanjeno punjenje EV (limit uvoza)');
	END_IF;
	IF xExpCurt AND NOT xPrevCurt THEN
		F_AlarmPush(k := kNow, sStamp := Team_HMI.sDateTime, iCode := 7, sText := 'Zastita prikljucka: ogranicena FNE (limit izvoza)');
	END_IF;
	IF xImpFail AND NOT xPrevFail THEN
		F_AlarmPush(k := kNow, sStamp := Team_HMI.sDateTime, iCode := 8, sText := 'UPOZORENJE: predvideni uvoz iznad limita');
	END_IF;
	xPrevShed := xEvShed;
	xPrevCurt := xExpCurt;
	xPrevFail := xImpFail;
	// remember for next step
	rGridPredLast := rGridPred;
	xHavePred := kNow < Team_Cfg.N_STEPS;
	FOR j := 0 TO 3 DO
		aPrevConn[j] := stOut.EV[j].connected AND kNow < Team_Cfg.N_STEPS;
		aPrevRemain[j] := stOut.EV[j].energy_required;
		aPrevDepK[j] := kNow + aEvSteps[j];
	END_FOR;
END_IF;

// ---------------- simulation state messages (every call, edge detected) ----------------
Team_HMI.xAlmTripped := stOut.sim_tripped OR SimCtrl.tripped;
Team_HMI.xAlmFinished := stOut.sim_finished OR SimCtrl.finished;
IF Team_HMI.xAlmTripped AND NOT xPrevTrip THEN
	F_AlarmPush(k := kNow, sStamp := Team_HMI.sDateTime, iCode := 3, sText := 'ODSPAJANJE od mreze (tripped) - simulacija zaustavljena');
END_IF;
IF Team_HMI.xAlmFinished AND NOT xPrevFin THEN
	F_AlarmPush(k := kNow, sStamp := Team_HMI.sDateTime, iCode := 4, sText := 'Simulacija godine zavrsena (finished)');
END_IF;
xPrevTrip := Team_HMI.xAlmTripped;
xPrevFin := Team_HMI.xAlmFinished;

(* ---- FB_Planner.st ---- *)
FUNCTION_BLOCK FB_Planner
// Rolling-horizon battery planner, re-solved every step (model predictive control).
//  1. Monthly peak cap T: the peak of the month so far is already paid, so T >= that peak.
//     A bisection finds the lowest cap the battery can hold over the PESSIMISTIC forecast
//     (aNetHi); T = max(peak so far, that cap * margin).
//  2. Dynamic programming over the stored battery energy (0..1200 kWh in 40 kWh levels):
//     cost(i) = import*TS*(price+fee) - export*TS*0.9*price(>=0) + PEN*(pessimistic import above T),
//     terminal value of stored energy = mean import price * PLAN_TVF.
//  3. The first interval is optimised with continuous candidates and the exact current values.
// Output rPb: requested BESS power for interval k (+ discharge / - charge); FB_GridGuard checks it.
VAR_INPUT
	iH : INT;                           // horizon length (1..192)
	rSoc : REAL;                        // [%]
	rBcMax : REAL;                      // feasible charge [kW]
	rBdMax : REAL;                      // feasible discharge [kW]
	rPeakSoFar : REAL;                  // import peak of the current month so far [kW]
	xHiInDp : BOOL;                     // TRUE: peak penalty uses the pessimistic net load
END_VAR
VAR_IN_OUT
	aNet : ARRAY[0..191] OF REAL;       // forecast net load without battery [kW] (i = 0 is exact)
	aNetHi : ARRAY[0..191] OF REAL;     // pessimistic net load for the peak cap [kW]
	aCi : ARRAY[0..191] OF REAL;        // import cost price + grid fee [EUR/kWh]
	aCe : ARRAY[0..191] OF REAL;        // export value 0.9*price, >= 0 [EUR/kWh]
END_VAR
VAR_OUTPUT
	rPb : REAL;                         // requested battery power, + discharge / - charge
	rT : REAL;                          // free import level (cap) used [kW]
	rTh : REAL;                         // cap under the pessimistic forecast [kW]
END_VAR
VAR CONSTANT
	NS : INT := 30;                     // energy levels 0..NS: 1200 kWh / 30 = 40 kWh per level
	AMIN : INT := -4;                   // max discharge levels per step (750*0.25/0.95/40 = 4.9)
	AMAX : INT := 4;                    // max charge levels per step (750*0.25*0.95/40 = 4.5)
	N_FIRST : INT := 21;                  // first-step candidates
END_VAR
VAR
	V : ARRAY[0..30] OF REAL;           // value function at i+1
	Vn : ARRAY[0..30] OF REAL;          // value function at i
	aBus : ARRAY[-4..4] OF REAL;        // bus power of each action, + discharge
	aCa : ARRAY[-4..4] OF REAL;         // stage cost of each action
	h : INT;
	i : INT;
	iE : INT;
	a : INT;
	m : INT;
	rDE : REAL;
	rEuse : REAL;
	rE0 : REAL;
	rE : REAL;
	rTv : REAL;
	rG : REAL;
	rC : REAL;
	rBest : REAL;
	rV : REAL;
	rB : REAL;
	rX : REAL;
	rFr : REAL;
	iS0 : INT;
	aCand : ARRAY[0..22] OF REAL;
	nCand : INT;
	ts : REAL;
	etaC : REAL;
	etaD : REAL;
	limImp : REAL;
	limExp : REAL;
END_VAR
// ---IMPL---
ts := SimParam.TS_H;
etaC := SimParam.BESS_ETA_CHG;
etaD := SimParam.BESS_ETA_DCH;
limImp := SimParam.EGC_MAX_IMPORT - Team_Cfg.GRID_MARGIN_IMP;
limExp := SimParam.EGC_MAX_EXPORT - Team_Cfg.GRID_MARGIN_EXP;
rEuse := (SimParam.BESS_SOC_MAX - SimParam.BESS_SOC_MIN) / 100.0 * SimParam.BESS_CAPACITY;
rDE := rEuse / INT_TO_REAL(NS);
h := LIMIT(1, iH, 192);
rE0 := (rSoc - SimParam.BESS_SOC_MIN) / 100.0 * SimParam.BESS_CAPACITY;

// ---------------- 1. monthly import caps ----------------
// rTh: cap the battery can hold under the PESSIMISTIC forecast (reserve)
// rT : free import level. Without PLAN_TSPLIT rT = rTh; with it rT is the cap needed under the
//      EXPECTED forecast, so the DP never plans grid charging above what the load needs anyway.
rTh := F_PeakCap(h := h, rE0 := rE0, rFloor := rPeakSoFar, rLimImp := limImp, aLoad := aNetHi);
IF Team_Cfg.PLAN_TSPLIT THEN
	rT := F_PeakCap(h := h, rE0 := rE0, rFloor := rPeakSoFar, rLimImp := limImp, aLoad := aNet);
ELSE
	rT := rTh;
END_IF;

// ---------------- 2. DP backward over stored energy ----------------
rTv := 0.0;
FOR i := 0 TO h - 1 DO
	rTv := rTv + aCi[i];
END_FOR;
rTv := rTv / INT_TO_REAL(h) * Team_Cfg.PLAN_TVF;
FOR iE := 0 TO NS DO
	V[iE] := -INT_TO_REAL(iE) * rDE * rTv;
END_FOR;
FOR a := AMIN TO AMAX DO
	IF a > 0 THEN
		aBus[a] := -INT_TO_REAL(a) * rDE / (ts * etaC);
	ELSE
		aBus[a] := -INT_TO_REAL(a) * rDE * etaD / ts;
	END_IF;
END_FOR;
FOR i := h - 1 TO 1 BY -1 DO
	FOR a := AMIN TO AMAX DO
		IF NOT Team_Cfg.PLAN_TSPLIT THEN
			IF xHiInDp THEN
				rG := aNetHi[i] - aBus[a];
			ELSE
				rG := aNet[i] - aBus[a];
			END_IF;
			aCa[a] := F_StageCost(aNet[i] - aBus[a], rG, aCi[i], aCe[i], rT, limExp);
		ELSE
			aCa[a] := F_StageCost(aNet[i] - aBus[a], aNet[i] - aBus[a], aCi[i], aCe[i], rT, limExp);
			IF xHiInDp AND aNetHi[i] - aBus[a] > rTh THEN
				aCa[a] := aCa[a] + Team_Cfg.PLAN_PEN * (aNetHi[i] - aBus[a] - rTh);
			END_IF;
		END_IF;
	END_FOR;
	FOR iE := 0 TO NS DO
		rBest := 3.0E38;
		FOR a := MAX(AMIN, -iE) TO MIN(AMAX, NS - iE) DO
			rV := aCa[a] + V[iE + a];
			IF rV < rBest THEN
				rBest := rV;
			END_IF;
		END_FOR;
		Vn[iE] := rBest;
	END_FOR;
	V := Vn;
END_FOR;

// ---------------- 3. first interval: continuous candidates ----------------
nCand := 0;
FOR m := 0 TO N_FIRST - 1 DO
	aCand[nCand] := -rBcMax + (rBcMax + rBdMax) * INT_TO_REAL(m) / INT_TO_REAL(N_FIRST - 1);
	nCand := nCand + 1;
END_FOR;
IF aNet[0] > -rBcMax AND aNet[0] < rBdMax THEN
	aCand[nCand] := aNet[0];            // exact self-consumption (grid = 0)
	nCand := nCand + 1;
END_IF;
IF aNet[0] - rT > -rBcMax AND aNet[0] - rT < rBdMax THEN
	aCand[nCand] := aNet[0] - rT;       // import exactly at the cap
	nCand := nCand + 1;
END_IF;
rBest := 3.0E38;
rPb := 0.0;
FOR m := 0 TO nCand - 1 DO
	rB := aCand[m];
	IF rB < 0.0 THEN
		rE := rE0 - rB * ts * etaC;
	ELSE
		rE := rE0 - rB * ts / etaD;
	END_IF;
	IF h > 1 THEN
		rX := LIMIT(0.0, rE / rDE, INT_TO_REAL(NS));
		iS0 := REAL_TO_INT(rX);             // REAL_TO_INT rounds -> make it floor
		IF INT_TO_REAL(iS0) > rX THEN
			iS0 := iS0 - 1;
		END_IF;
		iS0 := LIMIT(0, iS0, NS - 1);
		rFr := rX - INT_TO_REAL(iS0);
		rV := V[iS0] * (1.0 - rFr) + V[iS0 + 1] * rFr;
	ELSE
		rV := -rE * rTv;
	END_IF;
	rC := F_StageCost(aNet[0] - rB, aNet[0] - rB, aCi[0], aCe[0], rT, limExp) + rV;
	IF rC < rBest THEN
		rBest := rC;
		rPb := rB;
	END_IF;
END_FOR;
// never plan an import above the cap if the battery can avoid it
IF aNet[0] - rPb > rT THEN
	rPb := MIN(rBdMax, aNet[0] - rT);
END_IF;

(* ---- FB_Strategy.st ---- *)
FUNCTION_BLOCK FB_Strategy
// Energy-management strategy: decides the REQUESTED setpoints for interval k.
// Called once per new step. FB_GridGuard afterwards enforces the grid limits.
//   iMode 0 = baseline from spec 2.6: no curtailment, EVs at max power,
//             BESS charges only from PV surplus and discharges on deficit.
//   iMode 1 = optimised: forecast (FB_Forecast) + rolling-horizon planner (FB_Planner) for the
//             battery: monthly peak shaving + tariff / day-ahead arbitrage + PV self-consumption;
//             PV curtailed when the day-ahead price is negative and we would export.
VAR_INPUT
	iMode : INT;                        // strategy selector
	xReset : BOOL;                      // k = 0
	k : DINT;                           // current step
	iQh : INT;                          // qh_of_day
	iWeekday : INT;                     // 1 = Mon .. 7 = Sun
	iMonth : INT;                       // 1..12
	xVt : BOOL;                         // high tariff in interval k
	iPriceMode : INT;                   // SimCtrl.price_mode
	rFec : REAL;                        // fixed consumption interval k [kW]
	rFneAvail : REAL;                   // available PV interval k [kW]
	rSoc : REAL;                        // [%]
	rBcMax : REAL;                      // feasible BESS charge [kW]
	rBdMax : REAL;                      // feasible BESS discharge [kW]
	aEvMax : ARRAY[0..3] OF REAL;       // feasible EV power [kW]
	aEvRem : ARRAY[0..3] OF REAL;       // EV remaining energy [kWh] (0 if not connected)
	aEvSteps : ARRAY[0..3] OF DINT;     // EV steps to departure
	rPeakSoFar : REAL;                  // import peak of this month so far [kW]
END_VAR
VAR_OUTPUT
	rPbReq : REAL;                      // BESS request, + discharge / - charge [kW]
	aEvReq : ARRAY[0..3] OF REAL;       // EV requests [kW]
	xCurtReq : BOOL;                    // voluntary curtailment request
	rCurtReq : REAL;                    // PV limit [kW]
	rPeakTarget : REAL;                 // import cap aimed for (info for HMI) [kW]
	iHorizon : INT;                     // planning horizon used [steps]
END_VAR
VAR
	fbForecast : FB_Forecast;
	fbPlanner : FB_Planner;
	aNet : ARRAY[0..191] OF REAL;       // forecast net load
	aNetHi : ARRAY[0..191] OF REAL;     // pessimistic net load
	aVtF : ARRAY[0..191] OF BOOL;       // forecast VT
	aCi : ARRAY[0..191] OF REAL;        // import price + fee
	aCe : ARRAY[0..191] OF REAL;        // export value
	j : INT;
	i : INT;
	kk : DINT;
	sumEv : REAL;
	rP : REAL;
	rP0 : REAL;
END_VAR
// ---IMPL---
sumEv := 0.0;
FOR j := 0 TO 3 DO
	aEvReq[j] := aEvMax[j];             // EVs: charge at maximum feasible power (EV energy has priority)
	sumEv := sumEv + aEvReq[j];
END_FOR;
xCurtReq := FALSE;
rCurtReq := 0.0;

IF iMode = 0 THEN
	// ---------------- baseline (spec 2.6) ----------------
	// net demand on the bus without the battery: + deficit -> discharge, - PV surplus -> charge
	rPbReq := rFec + sumEv - rFneAvail;
	rPeakTarget := SimParam.EGC_MAX_IMPORT;
	iHorizon := 0;
ELSE
	// ---------------- optimised ----------------
	// horizon: PLAN_H steps; with day-ahead prices optionally only as far as prices are published
	// (tomorrow's prices are known after 13:00 = qh 52)
	IF iPriceMode = 1 AND Team_Cfg.PLAN_DA_PUBLISHED THEN
		iHorizon := 96 - iQh;
		IF iQh >= 52 THEN
			iHorizon := iHorizon + 96;
		END_IF;
		iHorizon := MIN(iHorizon, Team_Cfg.PLAN_H);   // cap the computing load (no measurable gain beyond 24 h)
	ELSE
		iHorizon := Team_Cfg.PLAN_H;
	END_IF;
	iHorizon := DINT_TO_INT(MIN(INT_TO_DINT(iHorizon), Team_Cfg.N_STEPS - k));
	iHorizon := LIMIT(1, iHorizon, 192);

	fbForecast(xReset := xReset, xUpdate := TRUE, k := k, iQh := iQh, iWeekday := iWeekday,
		rFec := rFec, rPv := rFneAvail, xVt := xVt, aEvRem := aEvRem, aEvSteps := aEvSteps,
		iH := iHorizon, rKsig := SEL(iPriceMode = 1, Team_Cfg.FC_KSIG_TT, Team_Cfg.FC_KSIG_DA),
		aNet := aNet, aNetHi := aNetHi, aVtF := aVtF);

	// prices over the horizon (price lists from Team_Prices, grid fee from SimParam)
	FOR i := 0 TO iHorizon - 1 DO
		kk := k + i;
		IF i = 0 THEN
			rP := F_EnergyPrice(k := kk, iMonth := iMonth, xHigh := xVt, iMode := iPriceMode);
			rP0 := rP;
		ELSE
			rP := F_EnergyPrice(k := kk, iMonth := iMonth, xHigh := aVtF[i], iMode := iPriceMode);
		END_IF;
		IF aVtF[i] THEN
			aCi[i] := rP + SimParam.GRID_VT;
		ELSE
			aCi[i] := rP + SimParam.GRID_NT;
		END_IF;
		aCe[i] := MAX(0.0, rP * SimParam.EXPORT_FACTOR);
	END_FOR;

	fbPlanner(iH := iHorizon, rSoc := rSoc, rBcMax := rBcMax, rBdMax := rBdMax, rPeakSoFar := rPeakSoFar,
		xHiInDp := SEL(iPriceMode = 1, Team_Cfg.PLAN_HI_TT, Team_Cfg.PLAN_HI_DA),
		aNet := aNet, aNetHi := aNetHi, aCi := aCi, aCe := aCe);
	rPbReq := fbPlanner.rPb;
	rPeakTarget := fbPlanner.rT;

	// negative energy price: do not export (export would cost money) -> curtail PV to the bus demand
	IF rP0 < 0.0 AND (rFec + sumEv - rPbReq - rFneAvail) < 0.0 THEN
		xCurtReq := TRUE;
		rCurtReq := MAX(0.0, rFec + sumEv - rPbReq);
	END_IF;
END_IF;

(* ---- Team_Main.st ---- *)
FUNCTION_BLOCK Team_Main
VAR_INPUT
      simOut : typeSimOut;
END_VAR
VAR_OUTPUT
      simCmd : typeSimCmd;
END_VAR
VAR_TEMP

END_VAR
VAR
	// ---- step sequencing (no timers: everything keyed on the simulated step k) ----
	xInit : BOOL;                       // first call done
	xNewStep : BOOL;                    // this call starts a new simulation step
	xResetStep : BOOL;                  // new step with k = 0 -> clear logs and state
	xLogNow : BOOL;                     // interval k-1 is logged in this step
	xHavePrev : BOOL;                   // values of interval k-1 are remembered
	kLast : DINT;                       // k of the previous new step
	dtLast : DT;                        // stamp of the previous new step
	k : DINT;
	j : INT;
	// ---- values of interval k-1 remembered for logging (spec 4.2) ----
	rFecPrev : REAL;                    // FEC_P_fix of interval k-1 (remembered for the next step)
	rFecLast : REAL;                    // FEC of the interval logged in this step (for HMI trend)
	iDayPrev : INT;                     // day_of_year of interval k-1
	iMonthPrev : INT;                   // month of interval k-1
	xHighPrev : BOOL;                   // VT of interval k-1
	aEvCmdPrev : ARRAY[0..3] OF REAL;   // feasible EV power commanded for interval k-1
	aEvConnPrev : ARRAY[0..3] OF BOOL;  // EV connected in interval k-1
	aEvDepKPrev : ARRAY[0..3] OF DINT;  // departure step of the EV connected in k-1
	aEvLast : ARRAY[0..3] OF REAL;      // actual EV power of interval k-1 (see note in body)
	rPrice : REAL;                      // energy price interval k
	rPricePrev : REAL;                  // energy price interval k-1
	// ---- per-step inputs for the control ----
	rBcMax : REAL;                      // feasible BESS charge [kW]
	rBdMax : REAL;                      // feasible BESS discharge [kW]
	aEvMax : ARRAY[0..3] OF REAL;       // feasible EV power [kW]
	aEvSteps : ARRAY[0..3] OF DINT;     // 15-min steps until departure
	aEvSlack : ARRAY[0..3] OF REAL;     // steps left minus steps needed at full power
	aEvRem : ARRAY[0..3] OF REAL;       // EV remaining energy [kWh] (0 if not connected)
	rPeakMonth : REAL;                  // import peak of the current month so far [kW]
	// ---- function blocks ----
	fbEnergyLog : FB_EnergyLogger;      // task 2
	fbCostLog : FB_CostLogger;          // task 3
	fbStrategy : FB_Strategy;           // task 1: what we would like to do
	fbGuard : FB_GridGuard;             // task 1: grid-limit protection (always last)
	fbHmi : FB_HmiUpdate;               // task 4 support data
	iStrategy : INT := 1;               // 0 = baseline (spec 2.6), 1 = forecast + planner
	// ---- command ----
	stCmd : typeSimCmd;                 // command for the current interval (held between steps)
	stCmdZero : typeSimCmd;             // never written -> all FALSE / 0
END_VAR

// ---IMPL---
// =====================================================================================
// Team_Main - energy manager. Called once per simulator step (SR_Main_Sim, phase 2 of 3).
// All state changes happen only when a NEW step is detected (k or stamp changed), so the
// result is independent of the SR_Main_Sim period. Order:
//   1. detect new step / reset   2. log interval k-1 (energy, cost)
//   3. control: strategy -> grid guard -> simCmd   4. remember values for the next step
//   5. HMI data. simCmd is written completely in every call.
// =====================================================================================
k := simOut.t_sim.k;
xNewStep := (NOT xInit) OR (k <> kLast) OR (simOut.t_sim.stamp <> dtLast);

IF xNewStep THEN
	xInit := TRUE;
	xResetStep := (k = 0);
	IF xResetStep THEN
		xHavePrev := FALSE;
	END_IF;

	// ---------------- 2. logging of interval k-1 ----------------
	xLogNow := xHavePrev AND (k = kLast + 1);
	FOR j := 0 TO 3 DO
		// The simulator publishes P_charge_act = 0 for an EV that departs at step k although it
		// was charged in interval k-1 (Sim_Core clears evPact on departure). For that interval we
		// use our own command, which was already clamped to the simulator's feasible value.
		IF xLogNow AND aEvConnPrev[j] AND (k >= aEvDepKPrev[j]) THEN
			aEvLast[j] := aEvCmdPrev[j];
		ELSE
			aEvLast[j] := simOut.EV[j].P_charge_act;
		END_IF;
	END_FOR;
	rFecLast := rFecPrev;
	IF xLogNow THEN
		rPricePrev := F_EnergyPrice(k := k - 1, iMonth := iMonthPrev, xHigh := xHighPrev, iMode := SimCtrl.price_mode);
	END_IF;
	fbEnergyLog(xReset := xResetStep, xLog := xLogNow, iDay := iDayPrev, iMonth := iMonthPrev,
		rFne := simOut.FNE_P_act, rFec := rFecPrev,
		rChg := simOut.BESS_P_charge_act, rDch := simOut.BESS_P_discharge_act,
		aEv := aEvLast, rImp := simOut.EGC_P_import, rExp := simOut.EGC_P_export);
	fbCostLog(xReset := xResetStep, xLog := xLogNow, iDay := iDayPrev, iMonth := iMonthPrev,
		rImp := simOut.EGC_P_import, rExp := simOut.EGC_P_export, rPrice := rPricePrev, xHigh := xHighPrev);

	// ---------------- 3. control ----------------
	IF (k >= Team_Cfg.N_STEPS) OR simOut.sim_finished THEN
		// final call (k = 35040): only logging, commands are ignored -> all zero
		stCmd := stCmdZero;
		xHavePrev := FALSE;
		FOR j := 0 TO 3 DO
			aEvCmdPrev[j] := 0.0;
			aEvConnPrev[j] := FALSE;
		END_FOR;
	ELSE
		rPrice := F_EnergyPrice(k := k, iMonth := simOut.t_sim.month, xHigh := simOut.t_sim.tariff_high, iMode := SimCtrl.price_mode);
		rPeakMonth := LREAL_TO_REAL(Team_Log.aMonth[LIMIT(1, simOut.t_sim.month, 12)].P_peak);
		// feasible limits (same clamps as the simulator)
		rBcMax := F_BessMaxChg(simOut.BESS_SoC);
		rBdMax := F_BessMaxDch(simOut.BESS_SoC);
		FOR j := 0 TO 3 DO
			IF simOut.EV[j].connected THEN
				aEvMax[j] := MAX(0.0, MIN(SimParam.EV_MAX_CHARGE,
					simOut.EV[j].energy_required / (SimParam.TS_H * SimParam.EV_ETA)));
				// planned departure is on a 15-min boundary: steps left = (departure - start of k) / 900 s
				aEvSteps[j] := MAX(1, (UDINT_TO_DINT(DT_TO_UDINT(simOut.EV[j].planned_departure))
					- UDINT_TO_DINT(DT_TO_UDINT(simOut.t_sim.stamp))) / 900);
				aEvSlack[j] := DINT_TO_REAL(aEvSteps[j])
					- simOut.EV[j].energy_required / (SimParam.EV_MAX_CHARGE * SimParam.TS_H * SimParam.EV_ETA);
				aEvRem[j] := simOut.EV[j].energy_required;
			ELSE
				aEvMax[j] := 0.0;
				aEvSteps[j] := 0;
				aEvSlack[j] := 0.0;
				aEvRem[j] := 0.0;
			END_IF;
		END_FOR;

		// 3a. strategy: requested setpoints
		fbStrategy(iMode := iStrategy, xReset := xResetStep, k := k, iQh := simOut.t_sim.qh_of_day,
			iWeekday := simOut.t_sim.weekday, iMonth := simOut.t_sim.month, xVt := simOut.t_sim.tariff_high,
			iPriceMode := SimCtrl.price_mode, rFec := simOut.FEC_P_fix, rFneAvail := simOut.FNE_output_power,
			rSoc := simOut.BESS_SoC, rBcMax := rBcMax, rBdMax := rBdMax, aEvMax := aEvMax,
			aEvRem := aEvRem, aEvSteps := aEvSteps, rPeakSoFar := rPeakMonth);

		// 3b. grid guard: predicted P_grid within EGC limits
		fbGuard(rFec := simOut.FEC_P_fix, rFneAvail := simOut.FNE_output_power,
			rBcMax := rBcMax, rBdMax := rBdMax, aEvMax := aEvMax, aEvSlack := aEvSlack,
			rPbReq := fbStrategy.rPbReq, aEvReq := fbStrategy.aEvReq,
			xCurtReq := fbStrategy.xCurtReq, rCurtReq := fbStrategy.rCurtReq);

		// 3c. complete command (all members, BESS enables mutually exclusive by construction)
		stCmd := stCmdZero;
		stCmd.FNE_enable_curtail := fbGuard.xCurt;
		stCmd.FNE_curtail_value := fbGuard.rCurt;
		IF fbGuard.rPb > Team_Cfg.P_EPS THEN
			stCmd.BESS_enable_discharge := TRUE;
			stCmd.BESS_P_discharge := fbGuard.rPb;
		ELSIF fbGuard.rPb < -Team_Cfg.P_EPS THEN
			stCmd.BESS_enable_charge := TRUE;
			stCmd.BESS_P_charge := -fbGuard.rPb;
		END_IF;
		FOR j := 0 TO 3 DO
			stCmd.EV[j].P_charge := fbGuard.aEv[j];
		END_FOR;

		// ---------------- 4. remember interval k for logging in step k+1 ----------------
		rFecPrev := simOut.FEC_P_fix;
		iDayPrev := simOut.t_sim.day_of_year;
		iMonthPrev := simOut.t_sim.month;
		xHighPrev := simOut.t_sim.tariff_high;
		FOR j := 0 TO 3 DO
			aEvCmdPrev[j] := fbGuard.aEv[j];
			aEvConnPrev[j] := simOut.EV[j].connected;
			aEvDepKPrev[j] := k + aEvSteps[j];
		END_FOR;
		xHavePrev := TRUE;
	END_IF;
	kLast := k;
	dtLast := simOut.t_sim.stamp;
END_IF;

// ---------------- 5. HMI data ----------------
fbHmi(xNewStep := xNewStep, xReset := xNewStep AND xResetStep, stOut := simOut, stCmd := stCmd,
	rPbCmd := fbGuard.rPb, rFneExp := fbGuard.rFne, rGridPred := fbGuard.rGridPred, rFecPrev := rFecLast,
	rPrice := rPrice, rPricePrev := rPricePrev, aEvSteps := aEvSteps, aEvLast := aEvLast,
	rPeakMonth := rPeakMonth, rPeakTarget := fbStrategy.rPeakTarget,
	xEvShed := fbGuard.xEvShed, xExpCurt := fbGuard.xExpCurt, xImpFail := fbGuard.xImpFail);

simCmd := stCmd;
